(* IEC 61131-3 sources: tree-sitter-st/tests/annexf, 13 files *)

(* ---- weigh.st ---- *)
FUNCTION WEIGH : WORD     (* BCD encoded *)
  VAR_INPUT  (* "EN" input is used to indicate "scale ready" *)
    weigh_command : BOOL;
    gross_weight : WORD ; (* BCD encoded *)
    tare_weight : INT ;
  END_VAR
(* Function Body *)
IF weigh_command THEN
  WEIGH := INT_TO_BCD (BCD_TO_INT(gross_weight) - tare_weight);
END_IF ;

END_FUNCTION                     (* Implicit "ENO" *)

(* ---- average.st ---- *)
 FUNCTION_BLOCK AVERAGE
   VAR_INPUT
     RUN : BOOL ;      (* 1 = run, 0 = reset *)
     XIN : REAL ;     (* Input variable *)
     N   : INT ;      (* 0 <= N < 128 or manufacturer- *)
   END_VAR            (*      specified maximum value  *)
   VAR_OUTPUT XOUT : REAL ; END_VAR (* Averaged output *)
   VAR SUM  : REAL := 0.0; (* Running sum *)
       FIFO : DELAY ;      (* N-Element FIFO *)
   END_VAR
   SUM := SUM - FIFO.XOUT ;
   FIFO (RUN := RUN , XIN := XIN, N := N) ;
   SUM := SUM + FIFO.XOUT ;
   IF RUN THEN XOUT := SUM/N ;
   ELSE SUM := N*XIN ; XOUT := XIN ;
   END_IF ;
 END_FUNCTION_BLOCK

(* ---- cmd_monitor.st ---- *)
FUNCTION_BLOCK CMD_MONITOR
 VAR_INPUT AUTO_CMD : BOOL ; (* Automated command *)
          AUTO_MODE : BOOL ; (* AUTO_CMD enable *)
            MAN_CMD : BOOL ; (* Manual Command *)
        MAN_CMD_CHK : BOOL ; (* Negated MAN_CMD to debounce *)
          T_CMD_MAX : TIME ; (* Max time from CMD to FDBK *)
               FDBK : BOOL ; (* Confirmation of CMD completion
                                by operative unit *)
                ACK : BOOL ; (* Acknowledge/cancel ALRM *)
 END_VAR
 VAR_OUTPUT CMD : BOOL ;   (* Command to operative unit *)
           ALRM : BOOL ;   (* T_CMD_MAX expired without FDBK *)
 END_VAR
 VAR
    CMD_TMR : TON ;    (* CMD-to-FDBK timer *)
    ALRM_FF : SR ;     (* Note over-riding S input: *)
 END_VAR                (* Command must be cancelled before
                              "ACK" can cancel alarm *)
    CMD := AUTO_CMD & AUTO_MODE
          OR MAN_CMD & NOT MAN_CMD_CHK & NOT AUTO_MODE ;

    CMD_TMR (IN := CMD, PT := T_CMD_MAX);
    ALRM_FF (S1 := CMD_TMR.Q & NOT FDBK, R := ACK);

    ALRM := ALRM_FF.Q1;
END_FUNCTION_BLOCK

(* ---- delay.st ---- *)
FUNCTION_BLOCK DELAY    (* N-sample delay *)
  VAR_INPUT
    RUN : BOOL ;     (* 1 = run, 0 = reset *)
    XIN : REAL ;
    N   : INT        (* 0 <= N < 128 or manufacturer- *)
  END_VAR            (*      specified maximum value  *)
  VAR_OUTPUT XOUT : REAL; END_VAR   (* Delayed output *)
  VAR X : ARRAY [0..127]     (* N-Element queue *)
               OF REAL;      (* with FIFO discipline *)
      I, IXIN, IXOUT : INT := 0;
  END_VAR
  IF RUN THEN
    IXIN := MOD(IXIN + 1, 128);
    X[IXIN] := XIN;
    IXOUT := MOD(IXOUT + 1, 128);
    XOUT := X[IXOUT];
  ELSE
    XOUT := XIN;
    IXIN := N;
    IXOUT := 0;
    FOR I := 0 TO N DO X[I] := XIN; END_FOR;
  END_IF ;
END_FUNCTION_BLOCK

(* ---- derivative.st ---- *)
 FUNCTION_BLOCK DERIVATIVE
   VAR_INPUT
     RUN : BOOL ;          (* 0 = reset                  *)
     XIN : REAL ;          (* Input to be differentiated *)
     CYCLE : TIME ;        (* Sampling period            *)
   END_VAR
   VAR_OUTPUT
     XOUT : REAL ;         (* Differentiated output      *)
   END_VAR
   VAR X1, X2, X3 : REAL ; END_VAR
   IF RUN THEN
      XOUT := (3.0 * (XIN - X3) + X1 - X2)
              / (10.0 * TIME_TO_REAL(CYCLE)) ;
      X3 := X2 ; X2 := X1 ; X1 := XIN ;
   ELSE XOUT := 0.0; X1 := XIN ; X2 := XIN ; X3 := XIN ;
   END_IF ;
 END_FUNCTION_BLOCK

(* ---- fwd_rev_mon.st ---- *)
FUNCTION_BLOCK FWD_REV_MON
VAR_INPUT AUTO : BOOL ;(* Enable automated commands *)
  ACK : BOOL ;         (* Acknowledge/cancel all alarms *)
  AUTO_FWD : BOOL ;    (* Automated forward command *)
  MAN_FWD : BOOL ;     (* Manual forward command *)
  MAN_FWD_CHK : BOOL ; (* Negated MAN_FWD for debouncing *)
  T_FWD_MAX : TIME ;  (* Maximum time from FWD_CMD to FWD_FDBK *)
  FWD_FDBK : BOOL ;    (* Confirmation of FWD_CMD completion *)
                       (*   by operative unit *)
  AUTO_REV : BOOL ;    (* Automated reverse command *)
  MAN_REV : BOOL ;     (* Manual reverse command *)
  MAN_REV_CHK : BOOL ; (* Negated MAN_REV for debouncing *)
  T_REV_MAX : TIME ;  (* Maximum time from REV_CMD to REV_FDBK *)
  REV_FDBK : BOOL ;    (* Confirmation of REV_CMD completion *)
END_VAR                (*    by operative unit *)
VAR_OUTPUT KLAXON : BOOL ;      (* Any alarm active *)
  FWD_REV_ALRM : BOOL; (* Forward/reverse command conflict *)
  FWD_CMD : BOOL ;     (* "Forward" command to operative unit *)
  FWD_ALRM : BOOL ;    (* T_FWD_MAX expired without FWD_FDBK *)
  REV_CMD : BOOL ;     (* "Reverse" command to operative unit *)
  REV_ALRM : BOOL ;    (* T_REV_MAX expired without REV_FDBK *)
END_VAR
VAR FWD_MON : CMD_MONITOR; (* "Forward" command monitor *)
  REV_MON : CMD_MONITOR;   (* "Reverse" command monitor *)
  FWD_REV_FF : SR ;      (* Forward/Reverse contention latch *)
END_VAR
(* Function Block body *)
(* Evaluate internal function blocks *)
  FWD_MON    (AUTO_MODE   := AUTO,
              ACK         := ACK,
              AUTO_CMD    := AUTO_FWD,
              MAN_CMD     := MAN_FWD,
              MAN_CMD_CHK := MAN_FWD_CHK,
              T_CMD_MAX   := T_FWD_MAX,
              FDBK        := FWD_FDBK);
  REV_MON    (AUTO_MODE   := AUTO,
              ACK         := ACK,
              AUTO_CMD    := AUTO_REV,
              MAN_CMD     := MAN_REV,
              MAN_CMD_CHK := MAN_REV_CHK,
              T_CMD_MAX   := T_REV_MAX,
              FDBK        := REV_FDBK);
  FWD_REV_FF (S1 := FWD_MON.CMD & REV_MON.CMD, R := ACK);
(* Transfer data to outputs *)
  FWD_REV_ALRM := FWD_REV_FF.Q1;
  FWD_CMD := FWD_MON.CMD & NOT FWD_REV_ALRM;
  FWD_ALRM := FWD_MON.ALRM;
  REV_CMD := REV_MON.CMD & NOT FWD_REV_ALRM;
  REV_ALRM := REV_MON.ALRM;
  KLAXON := FWD_ALRM OR REV_ALRM OR FWD_REV_ALRM;

END_FUNCTION_BLOCK

(* ---- hysteresis.st ---- *)
FUNCTION_BLOCK HYSTERESIS
    (* Boolean hysteresis on difference *)
    (* of REAL inputs, XIN1 - XIN2      *)
  VAR_INPUT XIN1, XIN2, EPS : REAL; END_VAR
  VAR_OUTPUT Q : BOOL := 0; END_VAR
  IF Q THEN IF XIN1 < (XIN2 - EPS) THEN Q := 0; END_IF ;
  ELSIF XIN1 > (XIN2 + EPS) THEN Q := 1 ;
  END_IF ;
END_FUNCTION_BLOCK

(* ---- integral.st ---- *)
 FUNCTION_BLOCK INTEGRAL
   VAR_INPUT
     RUN : BOOL ;       (* 1 = integrate, 0 = hold *)
     R1 : BOOL ;        (* Overriding reset        *)
     XIN : REAL ;       (* Input variable          *)
     X0  : REAL ;       (* Initial value           *)
     CYCLE : TIME ;     (* Sampling period         *)
   END_VAR
   VAR_OUTPUT
     Q : BOOL ;         (* NOT R1                  *)
     XOUT : REAL ;      (* Integrated output       *)
   END_VAR
   Q := NOT R1 ;
   IF R1 THEN XOUT := X0 ;
   ELSIF RUN THEN XOUT := XOUT + XIN * TIME_TO_REAL(CYCLE);
   END_IF ;
 END_FUNCTION_BLOCK

(* ---- lag1.st ---- *)
 FUNCTION_BLOCK LAG1
   VAR_INPUT
     RUN : BOOL ;     (* 1 = run, 0 = reset *)
     XIN : REAL ;     (* Input variable *)
     TAU : TIME ;     (* Filter time constant *)
     CYCLE : TIME ;   (* Sampling time interval *)
   END_VAR
   VAR_OUTPUT XOUT : REAL ; END_VAR  (* Filtered output *)
   VAR K : REAL ;     (* Smoothing constant, 0.0<=K<1.0 *)
   END_VAR
   IF RUN THEN XOUT := XOUT + K * (XIN - XOUT) ;
   ELSE XOUT := XIN ;
        K := TIME_TO_REAL(CYCLE) / TIME_TO_REAL(CYCLE + TAU) ;
   END_IF ;
 END_FUNCTION_BLOCK

(* ---- pid.st ---- *)
 FUNCTION_BLOCK PID
   VAR_INPUT
     AUTO : BOOL ;        (* 0 - manual , 1 - automatic *)
     PV : REAL ;          (* Process variable *)
     SP : REAL ;          (* Set point *)
     X0 : REAL ;          (* Manual output adjustment - *)
                          (* Typically from transfer station *)
     KP : REAL ;          (* Proportionality constant *)
     TR : REAL ;          (* Reset time *)
     TD : REAL ;          (* Derivative time constant *)
     CYCLE : TIME ;       (* Sampling period *)
   END_VAR
   VAR_OUTPUT XOUT : REAL; END_VAR
   VAR ERROR : REAL ;        (* PV - SP *)
       ITERM : INTEGRAL ;    (* FB for integral term  *)
       DTERM : DERIVATIVE ;  (* FB for derivative term *)
   END_VAR
   ERROR := PV - SP ;
   (*** Adjust ITERM so that XOUT := X0 when AUTO = 0 ***)
   ITERM (RUN := AUTO, R1 := NOT AUTO, XIN := ERROR,
          X0 := TR * (X0 - ERROR), CYCLE := CYCLE) ;
   DTERM (RUN := AUTO, XIN := ERROR, CYCLE := CYCLE) ;
   XOUT := KP * (ERROR + ITERM.XOUT/TR + DTERM.XOUT*TD) ;
 END_FUNCTION_BLOCK

(* ---- ramp.st ---- *)
 FUNCTION_BLOCK RAMP
   VAR_INPUT
     RUN : BOOL ;      (* 0 - track X0, 1 - ramp to/track X1 *)
     X0,X1 : REAL ;
     TR : TIME ;       (* Ramp duration *)
     CYCLE : TIME ;    (* Sampling period *)
   END_VAR
   VAR_OUTPUT
     BUSY : BOOL ; (* BUSY = 1 during ramping period *)
     XOUT : REAL := 0.0 ;
   END_VAR
   VAR XI : REAL ;       (* Initial value *)
       T : TIME := T#0s; (* Elapsed time of ramp *)
   END_VAR
   BUSY := RUN ;
   IF RUN THEN
      IF T >= TR THEN BUSY := 0 ; XOUT := X1 ;
      ELSE XOUT := XI + (X1-XI) * TIME_TO_REAL(T)
                                / TIME_TO_REAL(TR) ;
           T := T + CYCLE ;
      END_IF ;
   ELSE XOUT := X0 ; XI := X0 ; T := t#0s ;
   END_IF ;
 END_FUNCTION_BLOCK

(* ---- stack_int.st ---- *)
FUNCTION_BLOCK STACK_INT
  VAR_INPUT PUSH, POP: BOOL R_EDGE; (* Basic stack operations *)
            R1 : BOOL ;          (* Over-riding reset *)
            IN : INT ;           (* Input to be pushed *)
            N  : INT ;           (* Maximum depth after reset *)
  END_VAR
  VAR_OUTPUT EMPTY : BOOL := 1 ;     (* Stack empty *)
             OFLO  : BOOL := 0 ;     (* Stack overflow *)
             OUT   : INT  := 0 ;     (* Top of stack data *)
  END_VAR
  VAR STK : ARRAY[0..127] OF INT; (* Internal stack *)
      NI : INT :=128  ;           (* Storage for N upon reset *)
      PTR : INT := -1 ;           (* Stack pointer *)
  END_VAR
    (* Function Block body *)
    IF R1 THEN
       OFLO := 0; EMPTY := 1; PTR := -1;
       NI := LIMIT (MN:=1,IN:=N,MX:=128); OUT := 0;
    ELSIF POP & NOT EMPTY THEN
       OFLO := 0; PTR := PTR-1; EMPTY := PTR < 0;
       IF EMPTY THEN OUT := 0;
       ELSE OUT := STK[PTR];
       END_IF ;
    ELSIF PUSH & NOT OFLO THEN
       EMPTY := 0; PTR := PTR+1; OFLO := (PTR = NI);
       IF NOT OFLO THEN OUT := IN ; STK[PTR] := IN;
       ELSE OUT := 0;
       END_IF ;
    END_IF ;

  END_FUNCTION_BLOCK

(* ---- transfer.st ---- *)
FUNCTION_BLOCK TRANSFER
 VAR_INPUT
   AUTO : BOOL ;     (* 1 - track X0, 0 - ramp or hold *)
   XIN : REAL ;      (* Typically from PID Function Block *)
   FAST_RATE, SLOW_RATE : REAL ; (* Up/down ramp slopes *)
   FAST_UP, SLOW_UP, (* Typically pushbuttons *)
   FAST_DOWN, SLOW_DOWN : BOOL;
   CYCLE : TIME ;    (* Sampling period *)
 END_VAR
 VAR_OUTPUT XOUT : REAL ; END_VAR
 VAR XFER_RAMP : INTEGRAL ;
     RAMP_RATE : REAL ;
 END_VAR
 RAMP_RATE := 0.0 ;
 IF NOT AUTO THEN
  IF FAST_UP THEN RAMP_RATE := FAST_RATE; END_IF;
  IF SLOW_UP THEN RAMP_RATE := RAMP_RATE + SLOW_RATE; END_IF;
  IF FAST_DOWN THEN RAMP_RATE := RAMP_RATE - FAST_RATE; END_IF;
  IF SLOW_DOWN THEN RAMP_RATE := RAMP_RATE - SLOW_RATE; END_IF;
 END_IF ;
 XFER_RAMP (RUN := 1, CYCLE := CYCLE, R1 := AUTO,
            XIN := RAMP_RATE, X0 := XIN) ;
 XOUT := XFER_RAMP.XOUT;
END_FUNCTION_BLOCK
